       CASE #statRequest OF
         1:
           #data.parameterPage0 := #statParameterPage0;
         2:
           #data.systemCommand := #statSystemCommand;
         10:
           #data.vendorName := #statVendorName;
         11:
           #data.vendorText := #statVendorText;
         12:
           #data.productName := #statProductName;
         13:
           #data.productID := #statProductID;
         17:
           #data.fwRevision := #statFWRevision;
         18:
           #data.appSpecificName := #statAppSpecName;
         20:
           #data.statistics := #statStatistics;
         23:
           #data.diagnostics := #statDiagnostics;
         27:
           #data.parameters := #statParameters;
         ELSE // all other data sets are not defined
           ;
       END_CASE;
     END_IF;

     #statDone := #instDevice.done;
   END_REGION

   REGION OUTPUTS
     #done := #instDevice.done;
     #busy := #instDevice.busy;
     #error := #instDevice.error;
     #status := #instDevice.status;
     #diagDeviceFB := #instDevice.diagnostics;
   END_REGION
END_FUNCTION_BLOCK

// folder: Device-specific blocks/SIRIUS/3UG48

FUNCTION_BLOCK "LIOLink_3UG481x"   // FB5140, SCL
TITLE = LIOLink_3UG481x / IO_LINK_3UG481x
{ S7_Optimized_Access := 'FALSE' }
AUTHOR : SIOS
FAMILY : LIOLink
VERSION : 3.0
// IO-Link Device FB for SIRIUS 3UG481x to use with S7-300/400 controllers! / IO-Link Geraete FB fuer SIRIUS 3UG481x zur Nutzung mit S7-1500!
   VAR_INPUT
      execute : Bool;   // Request to execute function / Auftrag starten (mit steigender Flanke)
      logicalAddr : DInt;   // Logical address of IO-Link master module (sub module for ET 200eco PN) / Logische EA-Adresse des IO-Link Master Moduls
      cap : Int := 227;   // Client Access Point; 0xB400 for ET 200eco PN, CM 8x IO-Link, else 0xE003 (227) / Client Access Point (CAP), Siemens IO-Link Master immer 227 dezimal
      readWrite : Bool;   // FALSE: read, TRUE: write / Lese-/Schreibzugriff: 0=Lesen, 1=Schreiben
      port : Int;   // Port of the IO-Link Master for the Device / Port des Geraetes am IO-Link Mastermodul
      parameterPage0 : Bool := FALSE;   // Read access on parameter page 0 / Lesen Parameter Page 0
      systemCommands : Bool := FALSE;   // Write system commands / Schreiben Systemkommandos
      vendorName : Bool := FALSE;   // Read vendor name / Lesen Herstellername
      vendorText : Bool := FALSE;   // Read vendor text / Lesen Herstellertext
      productName : Bool := FALSE;   // Read product name / Lesen Produktname
      productID : Bool := FALSE;   // Read product ID / Lesen Produkt ID
      hwRevision : Bool := FALSE;   // Read hardware revision / Lesen HW-Revision
      fwRevision : Bool := FALSE;   // Read firmware revision / Lesen FW-Revision
      appSpecificName : Bool := FALSE;   // Read/Write application specific name / Lesen/Schreiben des spezifischen Applikationsnamen
      diagnostics : Bool := FALSE;   // Read diagnostics / Lesen der Diagnose
      measurements : Bool := FALSE;   // Read measurements / Lesen der Messwerte
      parameters : Bool;   // Read/Write parameters / Lesen/Schreiben der Parameter
   END_VAR
   VAR_OUTPUT
      done : Bool;   // TRUE: Commanded functionality has been completed successfully / Gueltigkeit 0: Daten ungueltig ; 1: Daten gueltig
      busy : Bool;   // TRUE: FB is not finished and new output values can be expected / 0: Auftrag beendet 1: Auftrag in Bearbeitung
      error : Bool;   // TRUE: An error occurred during the execution of the FB / Fehler = 0: kein Fehler; 1: Funktionsabbruch mit Fehler
      status : Word;   // 16#0000 - 16#7FFF: Status of the FB, 16#8000 - 16#FFFF: Error identification / DP/ PNIO - Fehlerstatus ; ERROR = 1 - Kommunikationsfehler in Detail
      diagDeviceFB : "LIOLink_typeDiagnostics";   // Diagnostics information of LIOLink_Device / IO-Link - Fehlerstatus; ERROR = 1: IO-Link Fehler in Detail
   END_VAR
   VAR_IN_OUT
      data : "LIOLink_3UG481_typeAll";   // Data area, device specific (Data Type) / Ablage der Gerätedaten, gerätespezifisch (Datentyp in DB)
   END_VAR
   VAR
      instDevice : "LIOLink_Device";
      statRecordParam : Struct   // Parameters to read/write specific records / Datensatzparameter (geraetespezifisch)
         index : Array[0..28] of Int;   // Index of data set / Datensatzindex
         subindex : Array[0..28] of Int;   // Subindex of data sets / Datensatzsubindex
         length : Array[0..28] of Int;   // Length of data set / Datensatzlänge
      END_STRUCT;
      statRecord : Array[0..231] of Byte;   // Record buffer
      statParameterPage0 AT statRecord : "LIOLink_typeParameterPage0";
      statSystemCommands AT statRecord : Byte;
      statVendorName AT statRecord : String[11];
      statVendorText AT statRecord : String[64];
      statProductName AT statRecord : String[64];
      statProductID AT statRecord : String[14];
      statHWRevision AT statRecord : String[7];
      statFWRevision AT statRecord : String[7];
      statAppSpecName AT statRecord : String[32];
      statDiagnostics AT statRecord : "LIOLink_3UG481_typeDiag";
      statMeasurements AT statRecord : "LIOLink_3UG481_typeMeasure";
      statParameters AT statRecord : "LIOLink_3UG481_typeParam";   // Product family SIRIUS (0x60)
      statIndex : Int;   // Requested index
      statSubindex : Int;   // Requested subindex
      statRecordLen : Int;   // Length of record to be written
      statRequest : Int;   // Case of request (data set) / Aktueller Fall (anfgefragter Datensatz)
      statDoneOld : Bool;   // Last cycle's value of instDevice.done
   END_VAR
   VAR_TEMP
      tempIndex : Int;   // Loop index
      tempLen : Int;   // Length
   END_VAR
   VAR CONSTANT
      MODE_READ : Bool := FALSE;   // Mode to read data
      MODE_WRITE : Bool := TRUE;   // Mode to write data
      STATUS_IDLE : Word := 16#7000;   // Status: Idle
   END_VAR
   // statRecordParam.index[3] := 2;
   // statRecordParam.index[2] := 0;
   // statRecordParam.index[1] := 0;
   // statRecordParam.index[0] := 0;
   // statRecordParam.index[17] := 23;
   // statRecordParam.index[16] := 22;
   // statRecordParam.index[5] := 0;
   // statRecordParam.index[4] := 0;
   // statRecordParam.index[15] := 21;
   // statRecordParam.index[14] := 20;
   // statRecordParam.index[13] := 19;
   // statRecordParam.index[12] := 18;
   // statRecordParam.index[11] := 17;
   // statRecordParam.index[10] := 16;
   // statRecordParam.index[9] := 0;
   // statRecordParam.index[8] := 0;
   // statRecordParam.index[7] := 0;
   // statRecordParam.index[6] := 0;
   // statRecordParam.length[28] := 60;
   // statRecordParam.length[27] := 0;
   // statRecordParam.length[26] := 0;
   // statRecordParam.length[25] := 38;
   // statRecordParam.length[24] := 30;
   // statRecordParam.length[23] := 0;
   // statRecordParam.length[22] := 0;
   // statRecordParam.length[21] := 0;
   // statRecordParam.length[20] := 0;
   // statRecordParam.length[19] := 0;
   // statRecordParam.length[18] := 32;
   // statRecordParam.length[17] := 7;
   // statRecordParam.length[16] := 7;
   // statRecordParam.length[15] := 0;
   // statRecordParam.length[14] := 0;
   // statRecordParam.length[13] := 14;
   // statRecordParam.length[12] := 64;
   // statRecordParam.length[11] := 64;
   // statRecordParam.length[10] := 11;
   // statRecordParam.length[9] := 0;
   // statRecordParam.length[8] := 0;
   // statRecordParam.length[7] := 0;
   // statRecordParam.length[6] := 0;
   // statRecordParam.length[5] := 0;
   // statRecordParam.length[4] := 0;
   // statRecordParam.length[3] := 1;
   // statRecordParam.length[2] := 0;
   // statRecordParam.length[1] := 16;
   // statRecordParam.length[0] := 0;
   // statRecordParam.index[28] := 131;
   // statRecordParam.index[27] := 0;
   // statRecordParam.index[26] := 0;
   // statRecordParam.index[25] := 94;
   // statRecordParam.index[24] := 92;
   // statRecordParam.index[23] := 0;
   // statRecordParam.index[22] := 0;
   // statRecordParam.index[21] := 0;
   // statRecordParam.index[20] := 0;
   // statRecordParam.index[19] := 0;
   // statRecordParam.index[18] := 24;
BEGIN
   REGION BLOCK INFO HEADER
     //===============================================================================
     // Siemens / (c)Copyright 2020
     //-------------------------------------------------------------------------------
     // Title:            LIOLink_3UG481x
     // Function:         Capsule block to communicate with 3UG481x devices
     // Library:          LIOLink
     // Author:           Siemens Industry Online Support
     // Tested with:      CPU 317-2 PN/DP FW 3.2
     // Engineering:      TIA Portal V16
     // Restrictions:     --
     // Requirements:     --
     //-------------------------------------------------------------------------------
     // Change log table:
     // Version  | Date       | Expert in charge       | Changes applied
     //----------|------------|------------------------|------------------------------
     // 01.00.00 | 11.04.2014 | Online Support         | First release
     // 01.01.00 | 12.09.2014 | Online Support         | Bugfixing write case 28 (data set 131)
     // 02.00.00 | 30.03.2015 | Online Support         | Upgrade to TIA Portal V13 SP1, use function IO_LINK_DEVICE, only one function for S7-1200 and 1500
     // 02.01.00 | 23.10.2015 | Online Support         | Upgraded FB "IO_LINK_DEVICE to V3.1.0
     // 03.00.00 | 22.09.2020 | Online Support         | Rewrote block for FB "LIOLink_Device" V4.0.0
     //===============================================================================
   END_REGION

   REGION INIT
     IF (#execute = TRUE AND #instDevice.status = #STATUS_IDLE) THEN
       // Request selector
       IF #parameterPage0 THEN
         #statRequest := 1;
       ELSIF #systemCommands THEN
         #statRequest := 3;
       ELSIF #vendorName THEN
         #statRequest := 10;
       ELSIF #vendorText THEN
         #statRequest := 11;
       ELSIF #productName THEN
         #statRequest := 12;
       ELSIF #productID THEN
         #statRequest := 13;
       ELSIF #hwRevision THEN
         #statRequest := 16;
       ELSIF #fwRevision THEN
         #statRequest := 17;
       ELSIF #appSpecificName THEN
         #statRequest := 18;
       ELSIF #diagnostics THEN
         #statRequest := 24;
       ELSIF #measurements THEN
         #statRequest := 25;
       ELSIF #parameters THEN
         #statRequest := 28;
       ELSE
         #statRequest := 0;
       END_IF;

       // Set request specific parameters
       #statIndex := #statRecordParam.index[#statRequest];
       #statSubindex := #statRecordParam.subindex[#statRequest];
       #statRecordLen := #statRecordParam.length[#statRequest];

       IF #readWrite = #MODE_WRITE THEN
         REGION write
           CASE #statRequest OF
             3:
               #statSystemCommands := #data.systemCommands;
             18:
               #statAppSpecName := #data.appSpecificName; // copy text into writing data
               #tempLen := LEN(#statAppSpecName); // determine length of text

               // Shift chars in array to remove String header
               FOR #tempIndex := 0 TO #tempLen - 1 DO
                 #statRecord[#tempIndex] := #statRecord[#tempIndex + 2]; // move [2] to [0], [3] to [1] ... until end of String
               END_FOR;

               // Fill remaining characters with null
               FOR #tempIndex := #tempLen TO #statRecordLen - 1 DO
                 #statRecord[#tempIndex] := CHAR_TO_BYTE('$00');
               END_FOR;
             28:
               #statParameters := #data.parameters;
             ELSE // All other data sets are read only  
               ;
           END_CASE;
         END_REGION

       END_IF;
     END_IF;
   END_REGION

   REGION CALL
     #instDevice(execute     := #execute,
                 logicalAddr := #logicalAddr,
                 cap         := #cap,
                 readWrite        := #readWrite,
                 "port"      := #port,
                 index       := #statIndex,
                 subindex    := #statSubindex,
                 writeLen    := #statRecordLen,
                 timeout     := T#20s,
                 record      := #statRecord);
   END_REGION

   REGION READ
     // Copy data
     IF #instDevice.done = TRUE AND #statDoneOld = FALSE AND #readWrite = #MODE_READ THEN
       IF (#statRequest >= 10 AND #statRequest <= 18) THEN // Only applies for String parameters (case 10..18)
         // Shift all characters to add string header
         FOR #tempIndex := (#statRecordLen + 1) TO 2 BY -1 DO
           #statRecord[#tempIndex] := #statRecord[#tempIndex - 2];
         END_FOR;
         // Add String header
         #statRecord[0] := INT_TO_BYTE(#statRecordLen);
         #statRecord[1] := INT_TO_BYTE(#statRecordLen);
       END_IF;

       CASE #statRequest OF
         1:
           #data.parameterPage0 := #statParameterPage0;
         10:
           #data.vendorName := #statVendorName;
         11:
           #data.vendorText := #statVendorText;
         12:
           #data.productName := #statProductName;
         13:
           #data.productID := #statProductID;
         16:
           #data.hwRevision := #statHWRevision;
         17:
           #data.fwRevision := #statFWRevision;
         18:
           #data.appSpecificName := #statAppSpecName;
         24:
           #data.diagnostics := #statDiagnostics;
         25:
           #data.measuredValues := #statMeasurements;
         28:
           #data.parameters := #statParameters;
         ELSE // Other data sets are not defined
           ;
       END_CASE;
     END_IF;

     #statDoneOld := #instDevice.done;
   END_REGION

   REGION OUTPUTS
     #done := #instDevice.done;
     #busy := #instDevice.busy;
     #error := #instDevice.error;
     #status := #instDevice.status;
     #diagDeviceFB := #instDevice.diagnostics;
   END_REGION
END_FUNCTION_BLOCK

FUNCTION_BLOCK "LIOLink_3UG4822"   // FB5150, SCL
TITLE = LIOLink_3UG4822 / IO_LINK_3UG4822_1500
{ S7_Optimized_Access := 'FALSE' }
AUTHOR : SIOS
FAMILY : LIOLink
VERSION : 3.0
// IO-Link Device FB for SIRIUS 3UG4822 to use with S7-300/400 controllers! / IO-Link Geraete FB fuer SIRIUS 3UG4822 zur Nutzung mit S7-1500!
   VAR_INPUT
      execute : Bool;   // Request to execute function / Auftrag starten (mit steigender Flanke)
      logicalAddr : DInt;   // Logical address of IO-Link master module (sub module for ET 200eco PN) / Logische EA-Adresse des IO-Link Master Moduls
      cap : Int := 227;   // Client Access Point; 0xB400 for ET 200eco PN, CM 8x IO-Link, else 0xE003 (227) / Client Access Point (CAP), Siemens IO-Link Master immer 227 dezimal
      readWrite : Bool;   // FALSE: read, TRUE: write / Lese-/Schreibzugriff: 0=Lesen, 1=Schreiben
      port : Int;   // Port of the IO-Link Master for the Device / Port des Geraetes am IO-Link Mastermodul
      parameterPage0 : Bool;   // Read access on parameter page 0 / Lesen Parameter Page 0
      systemCommands : Bool;   // Write system commands / Schreiben Systemkommandos
      vendorName : Bool;   // Read vendor name / Lesen Herstellername
      vendorText : Bool;   // Read vendor text / Lesen Herstellertext
      productName : Bool;   // Read product name / Lesen Produktname
      productID : Bool;   // Read product ID / Lesen Produkt ID
      hwRevision : Bool;   // Read hardware revision / Lesen HW-Revision
      fwRevision : Bool;   // Read firmware revision / Lesen FW-Revision
      appSpecificName : Bool;   // Read/Write application specific name / Lesen/Schreiben des spezifischen Applikationsnamen
      diagnostics : Bool;   // Read diagnostics / Lesen der Diagnose
      measurements : Bool;   // Read measurements / Lesen der Messwerte
      parameters : Bool;   // Read/Write parameters / Lesen/Schreiben der Parameter
   END_VAR
   VAR_OUTPUT
      done : Bool;   // TRUE: Commanded functionality has been completed successfully / Gueltigkeit 0: Daten ungueltig ; 1: Daten gueltig
      busy : Bool;   // TRUE: FB is not finished and new output values can be expected / 0: Auftrag beendet 1: Auftrag in Bearbeitung
      error : Bool;   // TRUE: An error occurred during the execution of the FB / Fehler = 0: kein Fehler; 1: Funktionsabbruch mit Fehler
      status : Word;   // 16#0000 - 16#7FFF: Status of the FB, 16#8000 - 16#FFFF: Error identification / DP/ PNIO - Fehlerstatus ; ERROR = 1 - Kommunikationsfehler in Detail
      diagDeviceFB : "LIOLink_typeDiagnostics";   // Diagnostics information of LIOLink_Device / IO-Link - Fehlerstatus; ERROR = 1: IO-Link Fehler in Detail
   END_VAR
   VAR_IN_OUT
      data : "LIOLink_3UG4822_typeAll";   // Data area, device specific (Data Type) / Ablage der Gerätedaten, gerätespezifisch (Datentyp in DB)
   END_VAR
   VAR
      instDevice : "LIOLink_Device";
      statRecordParam : Struct   // Parameters to read/write specific records / Datensatzparameter (geraetespezifisch)
         index : Array[0..28] of Int;   // Index of data set / Datensatzindex
         subindex : Array[0..28] of Int;   // Subindex of data sets / Datensatzsubindex
         length : Array[0..28] of Int;   // Length of data set / Datensatzlänge
      END_STRUCT;
      statRecord : Array[0..231] of Byte;   // Record buffer
      statParameterPage0 AT statRecord : "LIOLink_typeParameterPage0";
      statVendorName AT statRecord : String[11];
      statVendorText AT statRecord : String[64];
      statProductName AT statRecord : String[64];
      statProductID AT statRecord : String[14];
      statHWRevision AT statRecord : String[7];
      statFWRevision AT statRecord : String[7];
      statAppSpecName AT statRecord : String[32];
      statDiagnostics AT statRecord : "LIOLink_3UG4822_typeDiag";
      statMeasurements AT statRecord : "LIOLink_3UG4822_typeMeasure";
      statParameters AT statRecord : "LIOLink_3UG4822_typeParam";   // Product family SIRIUS (0x60)
      statSystemCommands AT statRecord : Byte;
      statIndex : Int;   // Requested index
      statSubindex : Int;   // Requested subindex
      statRecordLen : Int;   // Length of record to be written
      statRequest : Int;   // Case of request (data set) / Aktueller Fall (anfgefragter Datensatz)
      statDoneOld : Bool;   // Last cycle's value of instDevice.done
   END_VAR
   VAR_TEMP
      tempIndex : Int;   // Loop index
      tempLen : Int;   // Length
   END_VAR
   VAR CONSTANT
      MODE_READ : Bool := FALSE;   // Mode to read data
      MODE_WRITE : Bool := TRUE;   // Mode to write data
      STATUS_IDLE : Word := 16#7000;   // Status: Idle
   END_VAR
   // statRecordParam.index[3] := 2;
   // statRecordParam.index[2] := 0;
   // statRecordParam.index[1] := 0;
   // statRecordParam.index[0] := 0;
   // statRecordParam.index[17] := 23;
   // statRecordParam.index[16] := 22;
   // statRecordParam.index[5] := 0;
   // statRecordParam.index[4] := 0;
   // statRecordParam.index[15] := 21;
   // statRecordParam.index[14] := 20;
   // statRecordParam.index[13] := 19;
   // statRecordParam.index[12] := 18;
   // statRecordParam.index[11] := 17;
   // statRecordParam.index[10] := 16;
   // statRecordParam.index[9] := 0;
   // statRecordParam.index[8] := 0;
   // statRecordParam.index[7] := 0;
   // statRecordParam.index[6] := 0;
   // statRecordParam.length[28] := 64;
   // statRecordParam.length[27] := 0;
   // statRecordParam.length[26] := 0;
   // statRecordParam.length[25] := 52;
   // statRecordParam.length[24] := 28;
   // statRecordParam.length[23] := 0;
   // statRecordParam.length[22] := 0;
   // statRecordParam.length[21] := 0;
   // statRecordParam.length[20] := 0;
   // statRecordParam.length[19] := 0;
   // statRecordParam.length[18] := 32;
   // statRecordParam.length[17] := 7;
   // statRecordParam.length[16] := 7;
   // statRecordParam.length[15] := 0;
   // statRecordParam.length[14] := 0;
   // statRecordParam.length[13] := 14;
   // statRecordParam.length[12] := 64;
   // statRecordParam.length[11] := 64;
   // statRecordParam.length[10] := 11;
   // statRecordParam.length[9] := 0;
   // statRecordParam.length[8] := 0;
   // statRecordParam.length[7] := 0;
   // statRecordParam.length[6] := 0;
   // statRecordParam.length[5] := 0;
   // statRecordParam.length[4] := 0;
   // statRecordParam.length[3] := 1;
   // statRecordParam.length[2] := 0;
   // statRecordParam.length[1] := 16;
   // statRecordParam.length[0] := 0;
   // statRecordParam.index[28] := 131;
   // statRecordParam.index[27] := 0;
   // statRecordParam.index[26] := 0;
   // statRecordParam.index[25] := 94;
   // statRecordParam.index[24] := 92;
   // statRecordParam.index[23] := 0;
   // statRecordParam.index[22] := 0;
   // statRecordParam.index[21] := 0;
   // statRecordParam.index[20] := 0;
   // statRecordParam.index[19] := 0;
   // statRecordParam.index[18] := 24;
BEGIN
   REGION BLOCK INFO HEADER
     //===============================================================================
     // Siemens / (c)Copyright 2020
     //-------------------------------------------------------------------------------
     // Title:            LIOLink_3UG4822
     // Function:         Capsule block to communicate with 3UG4822 devices
     // Library:          LIOLink
     // Author:           Siemens Industry Online Support
     // Tested with:      CPU 317-2 PN/DP FW 3.2
     // Engineering:      TIA Portal V16
     // Restrictions:     --
     // Requirements:     --
     //-------------------------------------------------------------------------------
     // Change log table:
     // Version  | Date       | Expert in charge       | Changes applied
     //----------|------------|------------------------|------------------------------
     // 01.00.00 | 11.04.2014 | Online Support         | First release
     // 01.01.00 | 12.09.2014 | Online Support         | Bugfixing write case 28 (data set 131)
     // 02.00.00 | 30.03.2015 | Online Support         | Upgrade to TIA Portal V13 SP1, use function IO_LINK_DEVICE, only one function for S7-1200 and 1500
     // 02.01.00 | 23.10.2015 | Online Support         | Upgraded FB "IO_LINK_DEVICE to V3.1.0
     // 03.00.00 | 22.09.2020 | Online Support         | Rewrote block for FB "LIOLink_Device" V4.0.0
     //===============================================================================
   END_REGION

   REGION INIT
     IF (#execute = TRUE AND #instDevice.status = #STATUS_IDLE) THEN
       // Request selector
       IF #parameterPage0 THEN
         #statRequest := 1;
       ELSIF #systemCommands THEN
         #statRequest := 3;
       ELSIF #vendorName THEN
         #statRequest := 10;
       ELSIF #vendorText THEN
         #statRequest := 11;
       ELSIF #productName THEN
         #statRequest := 12;
       ELSIF #productID THEN
         #statRequest := 13;
       ELSIF #hwRevision THEN
         #statRequest := 16;
       ELSIF #fwRevision THEN
         #statRequest := 17;
       ELSIF #appSpecificName THEN
         #statRequest := 18;
       ELSIF #diagnostics THEN
         #statRequest := 24;
       ELSIF #measurements THEN
         #statRequest := 25;
       ELSIF #parameters THEN
         #statRequest := 28;
       ELSE
         #statRequest := 0;
       END_IF;

       // Set request specific parameters
       #statIndex := #statRecordParam.index[#statRequest];
       #statSubindex := #statRecordParam.subindex[#statRequest];
       #statRecordLen := #statRecordParam.length[#statRequest];

       IF #readWrite = #MODE_WRITE THEN
         REGION write
           CASE #statRequest OF
             3:
               #statSystemCommands := #data.systemCommands;
             18:
               #statAppSpecName := #data.appSpecificName; // copy text into writing data
               #tempLen := LEN(#statAppSpecName); // determine length of text

               // Shift chars in array to remove String header
               FOR #tempIndex := 0 TO #tempLen - 1 DO
                 #statRecord[#tempIndex] := #statRecord[#tempIndex + 2]; // move [2] to [0], [3] to [1] ... until end of String
               END_FOR;

               // Fill remaining characters with null
               FOR #tempIndex := #tempLen TO #statRecordLen - 1 DO
                 #statRecord[#tempIndex] := CHAR_TO_BYTE('$00');
               END_FOR;
             28:
               #statParameters := #data.parameters;
             ELSE // All other data sets are read only  
               ;
           END_CASE;
         END_REGION

       END_IF;
     END_IF;
   END_REGION

   REGION CALL
     #instDevice(execute     := #execute,
                 logicalAddr := #logicalAddr,
                 cap         := #cap,
                 readWrite   := #readWrite,
                 "port"      := #port,
                 index       := #statIndex,
                 subindex    := #statSubindex,
                 writeLen    := #statRecordLen,
                 timeout     := T#20s,
                 record      := #statRecord);
   END_REGION

   REGION READ
     // Copy data
     IF #instDevice.done = TRUE AND #statDoneOld = FALSE AND #readWrite = #MODE_READ THEN
       IF (#statRequest >= 10 AND #statRequest <= 18) THEN // Only applies for String parameters (case 10..18)
         // Shift all characters to add string header
         FOR #tempIndex := (#statRecordLen + 1) TO 2 BY -1 DO
           #statRecord[#tempIndex] := #statRecord[#tempIndex - 2];
         END_FOR;
         // Add String header
         #statRecord[0] := INT_TO_BYTE(#statRecordLen);
         #statRecord[1] := INT_TO_BYTE(#statRecordLen);
       END_IF;

       CASE #statRequest OF
         1:
           #data.parameterPage0 := #statParameterPage0;
         10:
           #data.vendorName := #statVendorName;
         11:
           #data.vendorText := #statVendorText;
         12:
           #data.productName := #statProductName;
         13:
           #data.productID := #statProductID;
         16:
           #data.hwRevision := #statHWRevision;
         17:
           #data.fwRevision := #statFWRevision;
         18:
           #data.appSpecificName := #statAppSpecName;
         24:
           #data.diagnostics := #statDiagnostics;
         25:
           #data.measuredValues := #statMeasurements;
         28:
           #data.parameters := #statParameters;
         ELSE // Other data sets are not defined
           ;
       END_CASE;
     END_IF;

     #statDoneOld := #instDevice.done;
   END_REGION

   REGION OUTPUTS
     #done := #instDevice.done;
     #busy := #instDevice.busy;
     #error := #instDevice.error;
     #status := #instDevice.status;
     #diagDeviceFB := #instDevice.diagnostics;
   END_REGION
END_FUNCTION_BLOCK

FUNCTION_BLOCK "LIOLink_3UG4825"   // FB5160, SCL
TITLE = LIOLink_3UG4825 / IO_LINK_3UG4825_1500
{ S7_Optimized_Access := 'FALSE' }
AUTHOR : SIOS
FAMILY : LIOLink
VERSION : 3.0
// IO-Link Device FB for SIRIUS 3UG4825 to use with S7-300/400 controllers! / IO-Link Geraete FB fuer SIRIUS 3UG4825 zur Nutzung mit S7-1500!
   VAR_INPUT
      execute : Bool;   // Request to execute function / Auftrag starten (mit steigender Flanke)
      logicalAddr : DInt;   // Logical address of IO-Link master module (sub module for ET 200eco PN) / Logische EA-Adresse des IO-Link Master Moduls
      cap : Int := 227;   // Client Access Point; 0xB400 for ET 200eco PN, CM 8x IO-Link, else 0xE003 (227) / Client Access Point (CAP), Siemens IO-Link Master immer 227 dezimal
      readWrite : Bool;   // FALSE: read, TRUE: write / Lese-/Schreibzugriff: 0=Lesen, 1=Schreiben
      port : Int;   // Port of the IO-Link Master for the Device / Port des Geraetes am IO-Link Mastermodul
      parameterPage0 : Bool;   // Read access on parameter page 0 / Lesen Parameter Page 0
      systemCommands : Bool;   // Write system commands / Schreiben Systemkommandos
      vendorName : Bool;   // Read vendor name / Lesen Herstellername
      vendorText : Bool;   // Read vendor text / Lesen Herstellertext
      productName : Bool;   // Read product name / Lesen Produktname
      productID : Bool;   // Read product ID / Lesen Produkt ID
      serialNumber : Bool;   // Read serial number / Lesen Seriennummer
      hwRevision : Bool;   // Read hardware revision / Lesen HW-Revision
      fwRevision : Bool;   // Read firmware revision / Lesen FW-Revision
      appSpecificName : Bool;   // Read/Write application specific name / Lesen/Schreiben des spezifischen Applikationsnamen
      diagnostics : Bool;   // Read diagnostics / Lesen der Diagnose
      measurements : Bool;   // Read measurements / Lesen der Messwerte
      parameters : Bool;   // Read/Write parameters / Lesen/Schreiben der Parameter
   END_VAR
   VAR_OUTPUT
      done : Bool;   // TRUE: Commanded functionality has been completed successfully / Gueltigkeit 0: Daten ungueltig ; 1: Daten gueltig
      busy : Bool;   // TRUE: FB is not finished and new output values can be expected / 0: Auftrag beendet 1: Auftrag in Bearbeitung
      error : Bool;   // TRUE: An error occurred during the execution of the FB / Fehler = 0: kein Fehler; 1: Funktionsabbruch mit Fehler
      status : Word;   // 16#0000 - 16#7FFF: Status of the FB, 16#8000 - 16#FFFF: Error identification / DP/ PNIO - Fehlerstatus ; ERROR = 1 - Kommunikationsfehler in Detail
      diagDeviceFB : "LIOLink_typeDiagnostics";   // Diagnostics information of LIOLink_Device / IO-Link - Fehlerstatus; ERROR = 1: IO-Link Fehler in Detail
   END_VAR
   VAR_IN_OUT
      data : "LIOLink_3UG4825_typeAll";   // Data area, device specific (Data Type) / Ablage der Gerätedaten, gerätespezifisch (Datentyp in DB)
   END_VAR
   VAR
      instDevice : "LIOLink_Device";
      statRecordParam : Struct   // Parameters to read/write specific records / Datensatzparameter (geraetespezifisch)
         index : Array[0..28] of Int;   // Index of data set / Datensatzindex
         subindex : Array[0..28] of Int;   // Subindex of data sets / Datensatzsubindex
         length : Array[0..28] of Int;   // Length of data set / Datensatzlänge
      END_STRUCT;
      statRecord : Array[0..231] of Byte;   // Record buffer
      statParameterPage0 AT statRecord : "LIOLink_typeParameterPage0";
      statVendorName AT statRecord : String[11];
      statVendorText AT statRecord : String[64];
      statProductName AT statRecord : String[64];
      statProductID AT statRecord : String[14];
      statSerialNumber AT statRecord : String[16];
      statHWRevision AT statRecord : String[7];
      statFWRevision AT statRecord : String[7];
      statAppSpecName AT statRecord : String[32];
      statDiagnostics AT statRecord : "LIOLink_3UG4825_typeDiag";
      statMeasurements AT statRecord : "LIOLink_3UG4825_typeMeasure";
      statParameters AT statRecord : "LIOLink_3UG4825_typeParam";   // Product family SIRIUS (0x60)
      statSystemCommands AT statRecord : Byte;
      statIndex : Int;   // Requested index
      statSubindex : Int;   // Requested subindex
      statRecordLen : Int;   // Length of record to be written
      statRequest : Int;   // Case of request (data set) / Aktueller Fall (anfgefragter Datensatz)
      statDoneOld : Bool;   // Last cycle's value of instDevice.done
   END_VAR
   VAR_TEMP
      tempIndex : Int;   // Loop index
      tempLen : Int;   // Length
   END_VAR
   VAR CONSTANT
      MODE_READ : Bool := FALSE;   // Mode to read data
      MODE_WRITE : Bool := TRUE;   // Mode to write data
      STATUS_IDLE : Word := 16#7000;   // Status: Idle
   END_VAR
   // statRecordParam.index[3] := 2;
   // statRecordParam.index[2] := 0;
   // statRecordParam.index[1] := 0;
   // statRecordParam.index[0] := 0;
   // statRecordParam.index[18] := 24;
   // statRecordParam.index[17] := 23;
   // statRecordParam.index[5] := 0;
   // statRecordParam.index[4] := 0;
   // statRecordParam.index[16] := 22;
   // statRecordParam.index[15] := 21;
   // statRecordParam.index[14] := 20;
   // statRecordParam.index[13] := 19;
   // statRecordParam.index[12] := 18;
   // statRecordParam.index[11] := 17;
   // statRecordParam.index[10] := 16;
   // statRecordParam.index[9] := 0;
   // statRecordParam.index[8] := 0;
   // statRecordParam.index[7] := 0;
   // statRecordParam.index[6] := 0;
   // statRecordParam.length[28] := 48;
   // statRecordParam.length[27] := 0;
   // statRecordParam.length[26] := 0;
   // statRecordParam.length[25] := 22;
   // statRecordParam.length[24] := 30;
   // statRecordParam.length[23] := 0;
   // statRecordParam.length[22] := 0;
   // statRecordParam.length[21] := 0;
   // statRecordParam.length[20] := 0;
   // statRecordParam.length[19] := 0;
   // statRecordParam.length[18] := 32;
   // statRecordParam.length[17] := 7;
   // statRecordParam.length[16] := 7;
   // statRecordParam.length[15] := 16;
   // statRecordParam.length[14] := 0;
   // statRecordParam.length[13] := 14;
   // statRecordParam.length[12] := 64;
   // statRecordParam.length[11] := 64;
   // statRecordParam.length[10] := 11;
   // statRecordParam.length[9] := 0;
   // statRecordParam.length[8] := 0;
   // statRecordParam.length[7] := 0;
   // statRecordParam.length[6] := 0;
   // statRecordParam.length[5] := 0;
   // statRecordParam.length[4] := 0;
   // statRecordParam.length[3] := 1;
   // statRecordParam.length[2] := 0;
   // statRecordParam.length[1] := 16;
   // statRecordParam.length[0] := 0;
   // statRecordParam.index[28] := 131;
   // statRecordParam.index[27] := 0;
   // statRecordParam.index[26] := 0;
   // statRecordParam.index[25] := 94;
   // statRecordParam.index[24] := 92;
   // statRecordParam.index[23] := 0;
   // statRecordParam.index[22] := 0;
   // statRecordParam.index[21] := 0;
   // statRecordParam.index[20] := 0;
   // statRecordParam.index[19] := 0;
BEGIN
   REGION BLOCK INFO HEADER
     //===============================================================================
     // Siemens / (c)Copyright 2020
     //-------------------------------------------------------------------------------
     // Title:            LIOLink_3UG4825
     // Function:         Capsule block to communicate with 3UG4825 devices
     // Library:          LIOLink
     // Author:           Siemens Industry Online Support
     // Tested with:      CPU 317-2 PN/DP FW 3.2
     // Engineering:      TIA Portal V16
     // Restrictions:     --
     // Requirements:     --
     //------------------------------------------------------------------------------
     // Change log table:
     // Version  | Date       | Expert in charge       | Changes applied
     //----------|------------|------------------------|------------------------------
     // 01.00.00 | 11.04.2014 | Online Support         | First release
     // 01.01.00 | 12.09.2014 | Online Support         | Bugfixing write case 28 (data set 131)
     // 02.00.00 | 30.03.2015 | Online Support         | Upgrade to TIA Portal V13 SP1, use function IO_LINK_DEVICE, only one function for S7-1200 and 1500
     // 02.01.00 | 23.10.2015 | Online Support         | Upgraded FB "IO_LINK_DEVICE to V3.1.0
     // 03.00.00 | 22.09.2020 | Online Support         | Rewrote block for FB "LIOLink_Device" V4.0.0
     //===============================================================================
   END_REGION

   REGION INIT
     IF (#execute = TRUE AND #instDevice.status = #STATUS_IDLE) THEN
       // Request selector
       IF #parameterPage0 THEN
         #statRequest := 1;
       ELSIF #systemCommands THEN
         #statRequest := 3;
       ELSIF #vendorName THEN
         #statRequest := 10;
       ELSIF #vendorText THEN
         #statRequest := 11;
       ELSIF #productName THEN
         #statRequest := 12;
       ELSIF #productID THEN
         #statRequest := 13;
       ELSIF #hwRevision THEN
         #statRequest := 16;
       ELSIF #fwRevision THEN
         #statRequest := 17;
       ELSIF #appSpecificName THEN
         #statRequest := 18;
       ELSIF #diagnostics THEN
         #statRequest := 24;
       ELSIF #measurements THEN
         #statRequest := 25;
       ELSIF #parameters THEN
         #statRequest := 28;
       ELSE
         #statRequest := 0;
       END_IF;

       // Set request specific parameters
       #statIndex := #statRecordParam.index[#statRequest];
       #statSubindex := #statRecordParam.subindex[#statRequest];
       #statRecordLen := #statRecordParam.length[#statRequest];

       IF #readWrite = #MODE_WRITE THEN
         REGION write
           CASE #statRequest OF
             3:
               #statSystemCommands := #data.systemCommands;
             18:
               #statAppSpecName := #data.appSpecificName; // copy text into writing data
               #tempLen := LEN(#statAppSpecName); // determine length of text

               // Shift chars in array to remove String header
               FOR #tempIndex := 0 TO #tempLen - 1 DO
                 #statRecord[#tempIndex] := #statRecord[#tempIndex + 2]; // move [2] to [0], [3] to [1] ... until end of String
               END_FOR;

               // Fill remaining characters with null
               FOR #tempIndex := #tempLen TO #statRecordLen - 1 DO
                 #statRecord[#tempIndex] := CHAR_TO_BYTE('$00');
               END_FOR;
             28:
               #statParameters := #data.parameters;
             ELSE // All other data sets are read only  
               ;
           END_CASE;
         END_REGION

       END_IF;
     END_IF;
   END_REGION

   REGION CALL
     #instDevice(execute     := #execute,
                 logicalAddr := #logicalAddr,
                 cap         := #cap,
                 readWrite   := #readWrite,
                 "port"      := #port,
                 index       := #statIndex,
                 subindex    := #statSubindex,
                 writeLen    := #statRecordLen,
                 timeout     := T#20s,
                 record      := #statRecord);
   END_REGION

   REGION READ
     // Copy data
     IF #instDevice.done = TRUE AND #statDoneOld = FALSE AND #readWrite = #MODE_READ THEN
       IF (#statRequest >= 10 AND #statRequest <= 18) THEN // Only applies for String parameters (case 10..18)
         // Shift all characters to add string header
         FOR #tempIndex := (#statRecordLen + 1) TO 2 BY -1 DO
           #statRecord[#tempIndex] := #statRecord[#tempIndex - 2];
         END_FOR;
         // Add String header
         #statRecord[0] := INT_TO_BYTE(#statRecordLen);
         #statRecord[1] := INT_TO_BYTE(#statRecordLen);
       END_IF;

       CASE #statRequest OF
         1:
           #data.parameterPage0 := #statParameterPage0;
         10:
           #data.vendorName := #statVendorName;
         11:
           #data.vendorText := #statVendorText;
         12:
           #data.productName := #statProductName;
         13:
           #data.productID := #statProductID;
         16:
           #data.hwRevision := #statHWRevision;
         17:
           #data.fwRevision := #statFWRevision;
         18:
           #data.appSpecificName := #statAppSpecName;
         24:
           #data.diagnostics := #statDiagnostics;
         25:
           #data.measuredValues := #statMeasurements;
         28:
           #data.parameters := #statParameters;
         ELSE // Other data sets are not defined
           ;
       END_CASE;
     END_IF;

     #statDoneOld := #instDevice.done;
   END_REGION

   REGION OUTPUTS
     #done := #instDevice.done;
     #busy := #instDevice.busy;
     #error := #instDevice.error;
     #status := #instDevice.status;
     #diagDeviceFB := #instDevice.diagnostics;
   END_REGION
END_FUNCTION_BLOCK

FUNCTION_BLOCK "LIOLink_3UG4832"   // FB5170, SCL
TITLE = LIOLink_3UG4832 / IO_LINK_3UG4832_1500
{ S7_Optimized_Access := 'FALSE' }
AUTHOR : SIOS
FAMILY : LIOLink
VERSION : 3.0
// IO-Link Device FB for SIRIUS 3UG4832 to use with S7-300/400 controllers! / IO-Link Geraete FB fuer SIRIUS 3UG4832 zur Nutzung mit S7-1500!
   VAR_INPUT
      execute : Bool;   // Request to execute function / Auftrag starten (mit steigender Flanke)
      logicalAddr : DInt;   // Logical address of IO-Link master module (sub module for ET 200eco PN) / Logische EA-Adresse des IO-Link Master Moduls
      cap : Int := 227;   // Client Access Point; 0xB400 for ET 200eco PN, CM 8x IO-Link, else 0xE003 (227) / Client Access Point (CAP), Siemens IO-Link Master immer 227 dezimal
      readWrite : Bool;   // FALSE: read, TRUE: write / Lese-/Schreibzugriff: 0=Lesen, 1=Schreiben
      port : Int;   // Port of the IO-Link Master for the Device / Port des Geraetes am IO-Link Mastermodul
      parameterPage0 : Bool;   // Read access on parameter page 0 / Lesen Parameter Page 0
      systemCommands : Bool;   // Write system commands / Schreiben Systemkommandos
      vendorName : Bool;   // Read vendor name / Lesen Herstellername
      vendorText : Bool;   // Read vendor text / Lesen Herstellertext
      productName : Bool;   // Read product name / Lesen Produktname
      productID : Bool;   // Read product ID / Lesen Produkt ID
      hwRevision : Bool;   // Read hardware revision / Lesen HW-Revision
      fwRevision : Bool;   // Read firmware revision / Lesen FW-Revision
      appSpecificName : Bool;   // Read/Write application specific name / Lesen/Schreiben des spezifischen Applikationsnamen
      diagnostics : Bool;   // Read diagnostics / Lesen der Diagnose
      measurements : Bool;   // Read measurements / Lesen der Messwerte
      parameters : Bool;   // Read/Write parameters / Lesen/Schreiben der Parameter
   END_VAR
   VAR_OUTPUT
      done : Bool;   // TRUE: Commanded functionality has been completed successfully / Gueltigkeit 0: Daten ungueltig ; 1: Daten gueltig
      busy : Bool;   // TRUE: FB is not finished and new output values can be expected / 0: Auftrag beendet 1: Auftrag in Bearbeitung
      error : Bool;   // TRUE: An error occurred during the execution of the FB / Fehler = 0: kein Fehler; 1: Funktionsabbruch mit Fehler
      status : Word;   // 16#0000 - 16#7FFF: Status of the FB, 16#8000 - 16#FFFF: Error identification / DP/ PNIO - Fehlerstatus ; ERROR = 1 - Kommunikationsfehler in Detail
      diagDeviceFB : "LIOLink_typeDiagnostics";   // Diagnostics information of LIOLink_Device / IO-Link - Fehlerstatus; ERROR = 1: IO-Link Fehler in Detail
   END_VAR
   VAR_IN_OUT
      data : "LIOLink_3UG4832_typeAll";   // Data area, device specific (Data Type) / Ablage der Gerätedaten, gerätespezifisch (Datentyp in DB)
   END_VAR
   VAR
      instDevice : "LIOLink_Device";
      statRecordParam : Struct   // Parameters to read/write specific records / Datensatzparameter (geraetespezifisch)
         index : Array[0..28] of Int;   // Index of data set / Datensatzindex
         subindex : Array[0..28] of Int;   // Subindex of data sets / Datensatzsubindex
         length : Array[0..28] of Int;   // Length of data set / Datensatzlänge
      END_STRUCT;
      statRecord : Array[0..231] of Byte;   // Record buffer
      statParameterPage0 AT statRecord : "LIOLink_typeParameterPage0";
      statVendorName AT statRecord : String[11];
      statVendorText AT statRecord : String[64];
      statProductName AT statRecord : String[64];
      statProductID AT statRecord : String[14];
      statHWRevision AT statRecord : String[7];
      statFWRevision AT statRecord : String[7];
      statAppSpecName AT statRecord : String[32];
      statDiagnostics AT statRecord : "LIOLink_3UG4832_typeDiag";
      statMeasurements AT statRecord : "LIOLink_3UG4832_typeMeasure";
      statParameters AT statRecord : "LIOLink_3UG4832_typeParam";   // Product family SIRIUS (0x60)
      statSystemCommands AT statRecord : Byte;
      statIndex : Int;   // Requested index
      statSubindex : Int;   // Requested subindex
      statRecordLen : Int;   // Length of record to be written
      statRequest : Int;   // Case of request (data set) / Aktueller Fall (anfgefragter Datensatz)
      statDoneOld : Bool;   // Last cycle's value of instDevice.done
   END_VAR
   VAR_TEMP
      tempIndex : Int;   // Loop index
      tempLen : Int;   // Length
   END_VAR
   VAR CONSTANT
      MODE_READ : Bool := FALSE;   // Mode to read data
      MODE_WRITE : Bool := TRUE;   // Mode to write data
      STATUS_IDLE : Word := 16#7000;   // Status: Idle
   END_VAR
   // statRecordParam.index[3] := 2;
   // statRecordParam.index[2] := 0;
   // statRecordParam.index[1] := 0;
   // statRecordParam.index[0] := 0;
   // statRecordParam.index[17] := 23;
   // statRecordParam.index[16] := 22;
   // statRecordParam.index[5] := 0;
   // statRecordParam.index[4] := 0;
   // statRecordParam.index[15] := 21;
   // statRecordParam.index[14] := 20;
   // statRecordParam.index[13] := 19;
   // statRecordParam.index[12] := 18;
   // statRecordParam.index[11] := 17;
   // statRecordParam.index[10] := 16;
   // statRecordParam.index[9] := 0;
   // statRecordParam.index[8] := 0;
   // statRecordParam.index[7] := 0;
   // statRecordParam.index[6] := 0;
   // statRecordParam.length[28] := 48;
   // statRecordParam.length[27] := 0;
   // statRecordParam.length[26] := 0;
   // statRecordParam.length[25] := 28;
   // statRecordParam.length[24] := 28;
   // statRecordParam.length[23] := 0;
   // statRecordParam.length[22] := 0;
   // statRecordParam.length[21] := 0;
   // statRecordParam.length[20] := 0;
   // statRecordParam.length[19] := 0;
   // statRecordParam.length[18] := 32;
   // statRecordParam.length[17] := 7;
   // statRecordParam.length[16] := 7;
   // statRecordParam.length[15] := 0;
   // statRecordParam.length[14] := 0;
   // statRecordParam.length[13] := 14;
   // statRecordParam.length[12] := 64;
   // statRecordParam.length[11] := 64;
   // statRecordParam.length[10] := 11;
   // statRecordParam.length[9] := 0;
   // statRecordParam.length[8] := 0;
   // statRecordParam.length[7] := 0;
   // statRecordParam.length[6] := 0;
   // statRecordParam.length[5] := 0;
   // statRecordParam.length[4] := 0;
   // statRecordParam.length[3] := 1;
   // statRecordParam.length[2] := 0;
   // statRecordParam.length[1] := 16;
   // statRecordParam.length[0] := 0;
   // statRecordParam.index[28] := 131;
   // statRecordParam.index[27] := 0;
   // statRecordParam.index[26] := 0;
   // statRecordParam.index[25] := 94;
   // statRecordParam.index[24] := 92;
   // statRecordParam.index[23] := 0;
   // statRecordParam.index[22] := 0;
   // statRecordParam.index[21] := 0;
   // statRecordParam.index[20] := 0;
   // statRecordParam.index[19] := 0;
   // statRecordParam.index[18] := 24;
BEGIN
   REGION BLOCK INFO HEADER
     //===============================================================================
     // Siemens / (c)Copyright 2020
     //-------------------------------------------------------------------------------
     // Title:            LIOLink_3UG4832
     // Function:         Capsule block to communicate with 3UG4832 devices
     // Library:          LIOLink
     // Author:           Siemens Industry Online Support
     // Tested with:      CPU 317-2 PN/DP FW 3.2
     // Engineering:      TIA Portal V16
     // Restrictions:     --
     // Requirements:     --
     //-------------------------------------------------------------------------------
     // Change log table:
     // Version  | Date       | Expert in charge       | Changes applied
     //----------|------------|------------------------|------------------------------
     // 01.00.00 | 11.04.2014 | Online Support         | First release
     // 01.01.00 | 12.09.2014 | Online Support         | Bugfixing write case 28 (data set 131)
     // 02.00.00 | 30.03.2015 | Online Support         | Upgrade to TIA Portal V13 SP1, use function IO_LINK_DEVICE, only one function for S7-1200 and 1500
     // 02.01.00 | 23.10.2015 | Online Support         | Upgraded FB "IO_LINK_DEVICE to V3.1.0
     // 03.00.00 | 22.09.2020 | Online Support         | Rewrote block for FB "LIOLink_Device" V4.0.0
     //===============================================================================
   END_REGION

   REGION INIT
     IF (#execute = TRUE AND #instDevice.status = #STATUS_IDLE) THEN
       // Request selector
       IF #parameterPage0 THEN
         #statRequest := 1;
       ELSIF #systemCommands THEN
         #statRequest := 3;
       ELSIF #vendorName THEN
         #statRequest := 10;
       ELSIF #vendorText THEN
         #statRequest := 11;
       ELSIF #productName THEN
         #statRequest := 12;
       ELSIF #productID THEN
         #statRequest := 13;
       ELSIF #hwRevision THEN
         #statRequest := 16;
       ELSIF #fwRevision THEN
         #statRequest := 17;
       ELSIF #appSpecificName THEN
         #statRequest := 18;
       ELSIF #diagnostics THEN
         #statRequest := 24;
       ELSIF #measurements THEN
         #statRequest := 25;
       ELSIF #parameters THEN
         #statRequest := 28;
       ELSE
         #statRequest := 0;
       END_IF;

       // Set request specific parameters
       #statIndex := #statRecordParam.index[#statRequest];
       #statSubindex := #statRecordParam.subindex[#statRequest];
       #statRecordLen := #statRecordParam.length[#statRequest];

       IF #readWrite = #MODE_WRITE THEN
         REGION write
           CASE #statRequest OF
             3:
               #statSystemCommands := #data.systemCommands;
             18:
               #statAppSpecName := #data.appSpecificName; // copy text into writing data
               #tempLen := LEN(#statAppSpecName); // determine length of text

               // Shift chars in array to remove String header
               FOR #tempIndex := 0 TO #tempLen - 1 DO
                 #statRecord[#tempIndex] := #statRecord[#tempIndex + 2]; // move [2] to [0], [3] to [1] ... until end of String
               END_FOR;

               // Fill remaining characters with null
               FOR #tempIndex := #tempLen TO #statRecordLen - 1 DO
                 #statRecord[#tempIndex] := CHAR_TO_BYTE('$00');
               END_FOR;
             28:
               #statParameters := #data.parameters;
             ELSE // All other data sets are read only  
               ;
           END_CASE;
         END_REGION

       END_IF;
     END_IF;
   END_REGION

   REGION CALL
     #instDevice(execute     := #execute,
                 logicalAddr := #logicalAddr,
                 cap         := #cap,
                 readWrite   := #readWrite,
                 "port"      := #port,
                 index       := #statIndex,
                 subindex    := #statSubindex,
                 writeLen    := #statRecordLen,
                 timeout     := T#20s,
                 record      := #statRecord);
   END_REGION

   REGION READ
     // Copy data
     IF #instDevice.done = TRUE AND #statDoneOld = FALSE AND #readWrite = #MODE_READ THEN
       IF (#statRequest >= 10 AND #statRequest <= 18) THEN // Only applies for String parameters (case 10..18)
         // Shift all characters to add string header
         FOR #tempIndex := (#statRecordLen + 1) TO 2 BY -1 DO
           #statRecord[#tempIndex] := #statRecord[#tempIndex - 2];
         END_FOR;
         // Add String header
         #statRecord[0] := INT_TO_BYTE(#statRecordLen);
         #statRecord[1] := INT_TO_BYTE(#statRecordLen);
       END_IF;

       CASE #statRequest OF
         1:
           #data.parameterPage0 := #statParameterPage0;
         10:
           #data.vendorName := #statVendorName;
         11:
           #data.vendorText := #statVendorText;
         12:
           #data.productName := #statProductName;
         13:
           #data.productID := #statProductID;
         16:
           #data.hwRevision := #statHWRevision;
         17:
           #data.fwRevision := #statFWRevision;
         18:
           #data.appSpecificName := #statAppSpecName;
         24:
           #data.diagnostics := #statDiagnostics;
         25:
           #data.measuredValues := #statMeasurements;
         28:
           #data.parameters := #statParameters;
         ELSE // Other data sets are not defined
           ;
       END_CASE;
     END_IF;

     #statDoneOld := #instDevice.done;
   END_REGION

   REGION OUTPUTS
     #done := #instDevice.done;
     #busy := #instDevice.busy;
     #error := #instDevice.error;
     #status := #instDevice.status;
     #diagDeviceFB := #instDevice.diagnostics;
   END_REGION
END_FUNCTION_BLOCK

FUNCTION_BLOCK "LIOLink_3UG4841"   // FB5180, SCL
TITLE = LIOLink_3UG4841 / IO_LINK_3UG4841_1500
{ S7_Optimized_Access := 'FALSE' }
AUTHOR : SIOS
FAMILY : LIOLink
VERSION : 3.0
// IO-Link Device FB for SIRIUS 3UG4841 to use with S7-300/400 controllers! / IO-Link Geraete FB fuer SIRIUS 3UG4841 zur Nutzung mit S7-1500!
   VAR_INPUT
      execute : Bool;   // Request to execute function / Auftrag starten (mit steigender Flanke)
      logicalAddr : DInt;   // Logical address of IO-Link master module (sub module for ET 200eco PN) / Logische EA-Adresse des IO-Link Master Moduls
      cap : Int := 227;   // Client Access Point; 0xB400 for ET 200eco PN, CM 8x IO-Link, else 0xE003 (227) / Client Access Point (CAP), Siemens IO-Link Master immer 227 dezimal
      readWrite : Bool;   // FALSE: read, TRUE: write / Lese-/Schreibzugriff: 0=Lesen, 1=Schreiben
      port : Int;   // Port of the IO-Link Master for the Device / Port des Geraetes am IO-Link Mastermodul
      parameterPage0 : Bool;   // Read access on parameter page 0 / Lesen Parameter Page 0
      systemCommands : Bool;   // Write system commands / Schreiben Systemkommandos
      vendorName : Bool;   // Read vendor name / Lesen Herstellername
      vendorText : Bool;   // Read vendor text / Lesen Herstellertext
      productName : Bool;   // Read product name / Lesen Produktname
      productID : Bool;   // Read product ID / Lesen Produkt ID
      hwRevision : Bool;   // Read hardware revision / Lesen HW-Revision
      fwRevision : Bool;   // Read firmware revision / Lesen FW-Revision
      appSpecificName : Bool;   // Read/Write application specific name / Lesen/Schreiben des spezifischen Applikationsnamen
      diagnostics : Bool;   // Read diagnostics / Lesen der Diagnose
      measurements : Bool;   // Read measurements / Lesen der Messwerte
      parameters : Bool;   // Read/Write parameters / Lesen/Schreiben der Parameter
   END_VAR
   VAR_OUTPUT
      done : Bool;   // TRUE: Commanded functionality has been completed successfully / Gueltigkeit 0: Daten ungueltig ; 1: Daten gueltig
      busy : Bool;   // TRUE: FB is not finished and new output values can be expected / 0: Auftrag beendet 1: Auftrag in Bearbeitung
      error : Bool;   // TRUE: An error occurred during the execution of the FB / Fehler = 0: kein Fehler; 1: Funktionsabbruch mit Fehler
      status : Word;   // 16#0000 - 16#7FFF: Status of the FB, 16#8000 - 16#FFFF: Error identification / DP/ PNIO - Fehlerstatus ; ERROR = 1 - Kommunikationsfehler in Detail
      diagDeviceFB : "LIOLink_typeDiagnostics";   // Diagnostics information of LIOLink_Device / IO-Link - Fehlerstatus; ERROR = 1: IO-Link Fehler in Detail
   END_VAR
   VAR_IN_OUT
      data : "LIOLink_3UG4841_typeAll";   // Data area, device specific (Data Type) / Ablage der Gerätedaten, gerätespezifisch (Datentyp in DB)
   END_VAR
   VAR
      instDevice : "LIOLink_Device";
      statRecordParam : Struct   // Parameters to read/write specific records / Datensatzparameter (geraetespezifisch)
         index : Array[0..28] of Int;   // Index of data set / Datensatzindex
         subindex : Array[0..28] of Int;   // Subindex of data sets / Datensatzsubindex
         length : Array[0..28] of Int;   // Length of data set / Datensatzlänge
      END_STRUCT;
      statRecord : Array[0..231] of Byte;   // Record buffer
      statParameterPage0 AT statRecord : "LIOLink_typeParameterPage0";
      statVendorName AT statRecord : String[11];
      statVendorText AT statRecord : String[64];
      statProductName AT statRecord : String[64];
      statProductID AT statRecord : String[14];
      statHWRevision AT statRecord : String[7];
      statFWRevision AT statRecord : String[7];
      statAppSpecName AT statRecord : String[32];
      statDiagnostics AT statRecord : "LIOLink_3UG4841_typeDiag";
      statMeasurements AT statRecord : "LIOLink_3UG4841_typeMeasure";
      statParameters AT statRecord : "LIOLink_3UG4841_typeParam";   // Product family SIRIUS (0x60)
      statSystemCommands AT statRecord : Byte;
      statIndex : Int;   // Requested index
      statSubindex : Int;   // Requested subindex
      statRecordLen : Int;   // Length of record to be written
      statRequest : Int;   // Case of request (data set) / Aktueller Fall (anfgefragter Datensatz)
      statDoneOld : Bool;   // Last cycle's value of instDevice.done
   END_VAR
   VAR_TEMP
      tempIndex : Int;   // Loop index
      tempLen : Int;   // Length
   END_VAR
   VAR CONSTANT
      MODE_READ : Bool := FALSE;   // Mode to read data
      MODE_WRITE : Bool := TRUE;   // Mode to write data
      STATUS_IDLE : Word := 16#7000;   // Status: Idle
   END_VAR
   // statRecordParam.index[3] := 2;
   // statRecordParam.index[2] := 0;
   // statRecordParam.index[1] := 0;
   // statRecordParam.index[0] := 0;
   // statRecordParam.index[17] := 23;
   // statRecordParam.index[16] := 22;
   // statRecordParam.index[5] := 0;
   // statRecordParam.index[4] := 0;
   // statRecordParam.index[15] := 21;
   // statRecordParam.index[14] := 20;
   // statRecordParam.index[13] := 19;
   // statRecordParam.index[12] := 18;
   // statRecordParam.index[11] := 17;
   // statRecordParam.index[10] := 16;
   // statRecordParam.index[9] := 0;
   // statRecordParam.index[8] := 0;
   // statRecordParam.index[7] := 0;
   // statRecordParam.index[6] := 0;
   // statRecordParam.length[28] := 74;
   // statRecordParam.length[27] := 0;
   // statRecordParam.length[26] := 0;
   // statRecordParam.length[25] := 50;
   // statRecordParam.length[24] := 30;
   // statRecordParam.length[23] := 0;
   // statRecordParam.length[22] := 0;
   // statRecordParam.length[21] := 0;
   // statRecordParam.length[20] := 0;
   // statRecordParam.length[19] := 0;
   // statRecordParam.length[18] := 32;
   // statRecordParam.length[17] := 7;
   // statRecordParam.length[16] := 7;
   // statRecordParam.length[15] := 0;
   // statRecordParam.length[14] := 0;
   // statRecordParam.length[13] := 14;
   // statRecordParam.length[12] := 64;
   // statRecordParam.length[11] := 64;
   // statRecordParam.length[10] := 11;
   // statRecordParam.length[9] := 0;
   // statRecordParam.length[8] := 0;
   // statRecordParam.length[7] := 0;
   // statRecordParam.length[6] := 0;
   // statRecordParam.length[5] := 0;
   // statRecordParam.length[4] := 0;
   // statRecordParam.length[3] := 1;
   // statRecordParam.length[2] := 0;
   // statRecordParam.length[1] := 16;
   // statRecordParam.length[0] := 0;
   // statRecordParam.index[28] := 131;
   // statRecordParam.index[27] := 0;
   // statRecordParam.index[26] := 0;
   // statRecordParam.index[25] := 94;
   // statRecordParam.index[24] := 92;
   // statRecordParam.index[23] := 0;
   // statRecordParam.index[22] := 0;
   // statRecordParam.index[21] := 0;
   // statRecordParam.index[20] := 0;
   // statRecordParam.index[19] := 0;
   // statRecordParam.index[18] := 24;
BEGIN
   REGION BLOCK INFO HEADER
     //===============================================================================
     // Siemens / (c)Copyright 2020
     //-------------------------------------------------------------------------------
     // Title:            LIOLink_3UG4841
     // Function:         Capsule block to communicate with 3UG4841 devices
     // Library:          LIOLink
     // Author:           Siemens Industry Online Support
     // Tested with:      CPU 317-2 PN/DP FW 3.2
     // Engineering:      TIA Portal V16
     // Restrictions:     --
     // Requirements:     --
     //-------------------------------------------------------------------------------
     // Change log table:
     // Version  | Date       | Expert in charge       | Changes applied
     //----------|------------|------------------------|------------------------------
     // 01.00.00 | 11.04.2014 | Online Support         | First release
     // 01.01.00 | 12.09.2014 | Online Support         | Bugfixing write case 28 (data set 131)
     // 02.00.00 | 30.03.2015 | Online Support         | Upgrade to TIA Portal V13 SP1, use function IO_LINK_DEVICE, only one function for S7-1200 and 1500
     // 02.01.00 | 23.10.2015 | Online Support         | Upgraded FB "IO_LINK_DEVICE to V3.1.0
     // 03.00.00 | 22.09.2020 | Online Support         | Rewrote block for FB "LIOLink_Device" V4.0.0
     //===============================================================================
   END_REGION

   REGION INIT
     IF (#execute = TRUE AND #instDevice.status = #STATUS_IDLE) THEN
       // Request selector
       IF #parameterPage0 THEN
         #statRequest := 1;
       ELSIF #systemCommands THEN
         #statRequest := 3;
       ELSIF #vendorName THEN
         #statRequest := 10;
       ELSIF #vendorText THEN
         #statRequest := 11;
       ELSIF #productName THEN
         #statRequest := 12;
       ELSIF #productID THEN
         #statRequest := 13;
       ELSIF #hwRevision THEN
         #statRequest := 16;
       ELSIF #fwRevision THEN
         #statRequest := 17;
       ELSIF #appSpecificName THEN
         #statRequest := 18;
       ELSIF #diagnostics THEN
         #statRequest := 24;
       ELSIF #measurements THEN
         #statRequest := 25;
       ELSIF #parameters THEN
         #statRequest := 28;
       ELSE
         #statRequest := 0;
       END_IF;

       // Set request specific parameters
       #statIndex := #statRecordParam.index[#statRequest];
       #statSubindex := #statRecordParam.subindex[#statRequest];
       #statRecordLen := #statRecordParam.length[#statRequest];

       IF #readWrite = #MODE_WRITE THEN
         REGION write
           CASE #statRequest OF
             3:
               #statSystemCommands := #data.systemCommands;
             18:
               #statAppSpecName := #data.appSpecificName; // copy text into writing data
               #tempLen := LEN(#statAppSpecName); // determine length of text

               // Shift chars in array to remove String header
               FOR #tempIndex := 0 TO #tempLen - 1 DO
                 #statRecord[#tempIndex] := #statRecord[#tempIndex + 2]; // move [2] to [0], [3] to [1] ... until end of String
               END_FOR;

               // Fill remaining characters with null
               FOR #tempIndex := #tempLen TO #statRecordLen - 1 DO
                 #statRecord[#tempIndex] := CHAR_TO_BYTE('$00');
               END_FOR;
             28:
               #statParameters := #data.parameters;
             ELSE // All other data sets are read only  
               ;
           END_CASE;
         END_REGION

       END_IF;
     END_IF;
   END_REGION

   REGION CALL
     #instDevice(execute     := #execute,
                 logicalAddr := #logicalAddr,
                 cap         := #cap,
                 readWrite   := #readWrite,
                 "port"      := #port,
                 index       := #statIndex,
                 subindex    := #statSubindex,
                 writeLen    := #statRecordLen,
                 timeout     := T#20s,
                 record      := #statRecord);
   END_REGION

   REGION READ
     // Copy data
     IF #instDevice.done = TRUE AND #statDoneOld = FALSE AND #readWrite = #MODE_READ THEN
       IF (#statRequest >= 10 AND #statRequest <= 18) THEN // Only applies for String parameters (case 10..18)
         // Shift all characters to add string header
         FOR #tempIndex := (#statRecordLen + 1) TO 2 BY -1 DO
           #statRecord[#tempIndex] := #statRecord[#tempIndex - 2];
         END_FOR;
         // Add String header
         #statRecord[0] := INT_TO_BYTE(#statRecordLen);
         #statRecord[1] := INT_TO_BYTE(#statRecordLen);
       END_IF;

       CASE #statRequest OF
         1:
           #data.parameterPage0 := #statParameterPage0;
         10:
           #data.vendorName := #statVendorName;
         11:
           #data.vendorText := #statVendorText;
         12:
           #data.productName := #statProductName;
         13:
           #data.productID := #statProductID;
         16:
           #data.hwRevision := #statHWRevision;
         17:
           #data.fwRevision := #statFWRevision;
         18:
           #data.appSpecificName := #statAppSpecName;
         24:
           #data.diagnostics := #statDiagnostics;
         25:
           #data.measuredValues := #statMeasurements;
         28:
           #data.parameters := #statParameters;
         ELSE // Other data sets are not defined
           ;
       END_CASE;
     END_IF;

     #statDoneOld := #instDevice.done;
   END_REGION

   REGION OUTPUTS
     #done := #instDevice.done;
     #busy := #instDevice.busy;
     #error := #instDevice.error;
     #status := #instDevice.status;
     #diagDeviceFB := #instDevice.diagnostics;
   END_REGION
END_FUNCTION_BLOCK

FUNCTION_BLOCK "LIOLink_3UG4851"   // FB5190, SCL
TITLE = LIOLink_3UG4851 / IO_LINK_3UG4851_1500
{ S7_Optimized_Access := 'FALSE' }
AUTHOR : SIOS
FAMILY : LIOLink
VERSION : 3.0
// IO-Link Device FB for SIRIUS 3UG4851 to use with S7-300/400 controllers! / IO-Link Geraete FB fuer SIRIUS 3UG4851 zur Nutzung mit S7-1500!
   VAR_INPUT
      execute : Bool;   // Request to execute function / Auftrag starten (mit steigender Flanke)
      logicalAddr : DInt;   // Logical address of IO-Link master module (sub module for ET 200eco PN) / Logische EA-Adresse des IO-Link Master Moduls
      cap : Int := 227;   // Client Access Point; 0xB400 for ET 200eco PN, CM 8x IO-Link, else 0xE003 (227) / Client Access Point (CAP), Siemens IO-Link Master immer 227 dezimal
      readWrite : Bool;   // FALSE: read, TRUE: write / Lese-/Schreibzugriff: 0=Lesen, 1=Schreiben
      port : Int;   // Port of the IO-Link Master for the Device / Port des Geraetes am IO-Link Mastermodul
      parameterPage0 : Bool;   // Read access on parameter page 0 / Lesen Parameter Page 0
      systemCommands : Bool;   // Write system commands / Schreiben Systemkommandos
      vendorName : Bool;   // Read vendor name / Lesen Herstellername
      vendorText : Bool;   // Read vendor text / Lesen Herstellertext
      productName : Bool;   // Read product name / Lesen Produktname
      productID : Bool;   // Read product ID / Lesen Produkt ID
      hwRevision : Bool;   // Read hardware revision / Lesen HW-Revision
      fwRevision : Bool;   // Read firmware revision / Lesen FW-Revision
      appSpecificName : Bool;   // Read/Write application specific name / Lesen/Schreiben des spezifischen Applikationsnamen
      diagnostics : Bool;   // Read diagnostics / Lesen der Diagnose
      measurements : Bool;   // Read measurements / Lesen der Messwerte
      parameters : Bool;   // Read/Write parameters / Lesen/Schreiben der Parameter
   END_VAR
   VAR_OUTPUT
      done : Bool;   // TRUE: Commanded functionality has been completed successfully / Gueltigkeit 0: Daten ungueltig ; 1: Daten gueltig
      busy : Bool;   // TRUE: FB is not finished and new output values can be expected / 0: Auftrag beendet 1: Auftrag in Bearbeitung
      error : Bool;   // TRUE: An error occurred during the execution of the FB / Fehler = 0: kein Fehler; 1: Funktionsabbruch mit Fehler
      status : Word;   // 16#0000 - 16#7FFF: Status of the FB, 16#8000 - 16#FFFF: Error identification / DP/ PNIO - Fehlerstatus ; ERROR = 1 - Kommunikationsfehler in Detail
      diagDeviceFB : "LIOLink_typeDiagnostics";   // Diagnostics information of LIOLink_Device / IO-Link - Fehlerstatus; ERROR = 1: IO-Link Fehler in Detail
   END_VAR
   VAR_IN_OUT
      data : "LIOLink_3UG4851_typeAll";   // Data area, device specific (Data Type) / Ablage der Gerätedaten, gerätespezifisch (Datentyp in DB)
   END_VAR
   VAR
      instDevice : "LIOLink_Device";
      statRecordParam : Struct   // Parameters to read/write specific records / Datensatzparameter (geraetespezifisch)
         index : Array[0..28] of Int;   // Index of data set / Datensatzindex
         subindex : Array[0..28] of Int;   // Subindex of data sets / Datensatzsubindex
         length : Array[0..28] of Int;   // Length of data set / Datensatzlänge
      END_STRUCT;
      statRecord : Array[0..231] of Byte;   // Record buffer
      statParameterPage0 AT statRecord : "LIOLink_typeParameterPage0";
      statVendorName AT statRecord : String[11];
      statVendorText AT statRecord : String[64];
      statProductName AT statRecord : String[64];
      statProductID AT statRecord : String[14];
      statHWRevision AT statRecord : String[7];
      statFWRevision AT statRecord : String[7];
      statAppSpecName AT statRecord : String[32];
      statDiagnostics AT statRecord : "LIOLink_3UG4851_typeDiag";
      statMeasurements AT statRecord : "LIOLink_3UG4851_typeMeasure";
      statParameters AT statRecord : "LIOLink_3UG4851_typeParam";   // Product family SIRIUS (0x60)
      statSystemCommands AT statRecord : Byte;
      statIndex : Int;   // Requested index
      statSubindex : Int;   // Requested subindex
      statRecordLen : Int;   // Length of record to be written
      statRequest : Int;   // Case of request (data set) / Aktueller Fall (anfgefragter Datensatz)
      statDoneOld : Bool;   // Last cycle's value of instDevice.done
   END_VAR
   VAR_TEMP
      tempIndex : Int;   // Loop index
      tempLen : Int;   // Length
   END_VAR
   VAR CONSTANT
      MODE_READ : Bool := FALSE;   // Mode to read data
      MODE_WRITE : Bool := TRUE;   // Mode to write data
      STATUS_IDLE : Word := 16#7000;   // Status: Idle
   END_VAR
   // statRecordParam.index[3] := 2;
   // statRecordParam.index[2] := 0;
   // statRecordParam.index[1] := 0;
   // statRecordParam.index[0] := 0;
   // statRecordParam.index[17] := 23;
   // statRecordParam.index[16] := 22;
   // statRecordParam.index[5] := 0;
   // statRecordParam.index[4] := 0;
   // statRecordParam.index[15] := 21;
   // statRecordParam.index[14] := 20;
   // statRecordParam.index[13] := 19;
   // statRecordParam.index[12] := 18;
   // statRecordParam.index[11] := 17;
   // statRecordParam.index[10] := 16;
   // statRecordParam.index[9] := 0;
   // statRecordParam.index[8] := 0;
   // statRecordParam.index[7] := 0;
   // statRecordParam.index[6] := 0;
   // statRecordParam.length[28] := 48;
   // statRecordParam.length[27] := 0;
   // statRecordParam.length[26] := 0;
   // statRecordParam.length[25] := 18;
   // statRecordParam.length[24] := 30;
   // statRecordParam.length[23] := 0;
   // statRecordParam.length[22] := 0;
   // statRecordParam.length[21] := 0;
   // statRecordParam.length[20] := 0;
   // statRecordParam.length[19] := 0;
   // statRecordParam.length[18] := 32;
   // statRecordParam.length[17] := 7;
   // statRecordParam.length[16] := 7;
   // statRecordParam.length[15] := 0;
   // statRecordParam.length[14] := 0;
   // statRecordParam.length[13] := 14;
   // statRecordParam.length[12] := 64;
   // statRecordParam.length[11] := 64;
   // statRecordParam.length[10] := 11;
   // statRecordParam.length[9] := 0;
   // statRecordParam.length[8] := 0;
   // statRecordParam.length[7] := 0;
   // statRecordParam.length[6] := 0;
   // statRecordParam.length[5] := 0;
   // statRecordParam.length[4] := 0;
   // statRecordParam.length[3] := 1;
   // statRecordParam.length[2] := 0;
   // statRecordParam.length[1] := 16;
   // statRecordParam.length[0] := 0;
   // statRecordParam.index[28] := 131;
   // statRecordParam.index[27] := 0;
   // statRecordParam.index[26] := 0;
   // statRecordParam.index[25] := 94;
   // statRecordParam.index[24] := 92;
   // statRecordParam.index[23] := 0;
   // statRecordParam.index[22] := 0;
   // statRecordParam.index[21] := 0;
   // statRecordParam.index[20] := 0;
   // statRecordParam.index[19] := 0;
   // statRecordParam.index[18] := 24;
BEGIN
   REGION BLOCK INFO HEADER
     //===============================================================================
     // Siemens / (c)Copyright 2020
     //-------------------------------------------------------------------------------
     // Title:            LIOLink_3UG4851
     // Function:         Capsule block to communicate with 3UG4851 devices
     // Library:          LIOLink
     // Author:           Siemens Industry Online Support
     // Tested with:      CPU 317-2 PN/DP FW 3.2
     // Engineering:      TIA Portal V16
     // Restrictions:     --
     // Requirements:     --
     //-------------------------------------------------------------------------------
     // Change log table:
     // Version  | Date       | Expert in charge       | Changes applied
     //----------|------------|------------------------|------------------------------
     // 01.00.00 | 11.04.2014 | Online Support         | First release
     // 01.01.00 | 12.09.2014 | Online Support         | Bugfixing write case 28 (data set 131)
     // 02.00.00 | 30.03.2015 | Online Support         | Upgrade to TIA Portal V13 SP1, use function IO_LINK_DEVICE, only one function for S7-1200 and 1500
     // 02.01.00 | 23.10.2015 | Online Support         | Upgraded FB "IO_LINK_DEVICE to V3.1.0
     // 03.00.00 | 22.09.2020 | Online Support         | Rewrote block for FB "LIOLink_Device" V4.0.0
     //===============================================================================
   END_REGION

   REGION INIT
     IF (#execute = TRUE AND #instDevice.status = #STATUS_IDLE) THEN
       // Request selector
       IF #parameterPage0 THEN
         #statRequest := 1;
       ELSIF #systemCommands THEN
         #statRequest := 3;
       ELSIF #vendorName THEN
         #statRequest := 10;
       ELSIF #vendorText THEN
         #statRequest := 11;
       ELSIF #productName THEN
         #statRequest := 12;
       ELSIF #productID THEN
         #statRequest := 13;
       ELSIF #hwRevision THEN
         #statRequest := 16;
       ELSIF #fwRevision THEN
         #statRequest := 17;
       ELSIF #appSpecificName THEN
         #statRequest := 18;
       ELSIF #diagnostics THEN
         #statRequest := 24;
       ELSIF #measurements THEN
         #statRequest := 25;
       ELSIF #parameters THEN
         #statRequest := 28;
       ELSE
         #statRequest := 0;
       END_IF;

       // Set request specific parameters
       #statIndex := #statRecordParam.index[#statRequest];
       #statSubindex := #statRecordParam.subindex[#statRequest];
       #statRecordLen := #statRecordParam.length[#statRequest];

       IF #readWrite = #MODE_WRITE THEN
         REGION write
           CASE #statRequest OF
             3:
               #statSystemCommands := #data.systemCommands;
             18:
               #statAppSpecName := #data.appSpecificName; // copy text into writing data
               #tempLen := LEN(#statAppSpecName); // determine length of text

               // Shift chars in array to remove String header
               FOR #tempIndex := 0 TO #tempLen - 1 DO
                 #statRecord[#tempIndex] := #statRecord[#tempIndex + 2]; // move [2] to [0], [3] to [1] ... until end of String
               END_FOR;

               // Fill remaining characters with null
               FOR #tempIndex := #tempLen TO #statRecordLen - 1 DO
                 #statRecord[#tempIndex] := CHAR_TO_BYTE('$00');
               END_FOR;
             28:
               #statParameters := #data.parameters;
             ELSE // All other data sets are read only  
               ;
           END_CASE;
         END_REGION

       END_IF;
     END_IF;
   END_REGION

   REGION CALL
     #instDevice(execute     := #execute,
                 logicalAddr := #logicalAddr,
                 cap         := #cap,
                 readWrite   := #readWrite,
                 "port"      := #port,
                 index       := #statIndex,
                 subindex    := #statSubindex,
                 writeLen    := #statRecordLen,
                 timeout     := T#20s,
                 record      := #statRecord);
   END_REGION

   REGION READ
     // Copy data
     IF #instDevice.done = TRUE AND #statDoneOld = FALSE AND #readWrite = #MODE_READ THEN
       IF (#statRequest >= 10 AND #statRequest <= 18) THEN // Only applies for String parameters (case 10..18)
         // Shift all characters to add string header
         FOR #tempIndex := (#statRecordLen + 1) TO 2 BY -1 DO
           #statRecord[#tempIndex] := #statRecord[#tempIndex - 2];
         END_FOR;
         // Add String header
         #statRecord[0] := INT_TO_BYTE(#statRecordLen);
         #statRecord[1] := INT_TO_BYTE(#statRecordLen);
       END_IF;

       CASE #statRequest OF
         1:
           #data.parameterPage0 := #statParameterPage0;
         10:
           #data.vendorName := #statVendorName;
         11:
           #data.vendorText := #statVendorText;
         12:
           #data.productName := #statProductName;
         13:
           #data.productID := #statProductID;
         16:
           #data.hwRevision := #statHWRevision;
         17:
           #data.fwRevision := #statFWRevision;
         18:
           #data.appSpecificName := #statAppSpecName;
         24:
           #data.diagnostics := #statDiagnostics;
         25:
           #data.measuredValues := #statMeasurements;
         28:
           #data.parameters := #statParameters;
         ELSE // Other data sets are not defined
           ;
       END_CASE;
     END_IF;

     #statDoneOld := #instDevice.done;
   END_REGION

   REGION OUTPUTS
     #done := #instDevice.done;
     #busy := #instDevice.busy;
     #error := #instDevice.error;
     #status := #instDevice.status;
     #diagDeviceFB := #instDevice.diagnostics;
   END_REGION
END_FUNCTION_BLOCK

// folder: Devices/SIMATIC RF200

FUNCTION_BLOCK "LIOLink_RF200_ReadTag"   // FB2, SCL
TITLE = LRfidIOL_Read
{ S7_Optimized_Access := 'FALSE' }
FAMILY : S7-300
VERSION : 3.1
// Read Data with IO-Link readers
// IO-Link V1.1
   VAR_INPUT
      execute : Bool;
      addrTag : Word;
      length : Word;
      hwID : Word;
      portAddr : Int;
      "version" : Int;
   END_VAR
   VAR_OUTPUT
      done : Bool;
      busy : Bool;
      error : Bool;
      status : DWord;
      statusWord AT status : Array[0..1] of Word;
      presence : Bool;
   END_VAR
   VAR_IN_OUT
      identData : ANY;
   END_VAR
   VAR
      statPae : Array[0..28] of Byte;
      Status_Byte : Byte;
      Status_bit AT Status_Byte : Array[0..7] of Bool;
      statPresence : Bool;
      statNState : Int;
      statIdleState : Int;
      statTelegramState : Int := 1;
      statReadState : Int := 2;
      statErrorState : Int := 3;
      statAdr : Word;
      statAdrRead AT statAdr : Array[0..1] of Byte;
      statBlk : Int;
      statReadOffset : Int := 0;
      statExecuteReq : Bool;
      statOffset : DInt;
      statOffset2 : DWord;
      statLength : DInt;
      statDat : Array[0..31] of Byte;
      statRecDat : Array[0..31] of Byte;
      statAddrOffset : Int;
      statPresenceFF : Bool;
      statTimerIn : Bool;
      statTimerPt : Time := T#5s;
      instTon : TON;
      statDone : Bool;
      statBusy : Bool;
      InstSetIoPart : SETIO_PART;
      statIoPartError : Bool;
      statIoPartStatus : DWord;
      InstGetIoPart : GETIO_PART;
      statIOsizeNetto : Int;
      statIOsize : Int;
   END_VAR
   VAR_TEMP
      tempSPointer : ANY;
      tempPoint1 AT tempSPointer : Struct
         dentifier : Byte;
         typ : Byte;
         length : Int;
         dbnr : Int;
         datapointer : DWord;
      END_STRUCT;
      tempDPointer : ANY;
      tempPoint2 AT tempDPointer : Struct
         dentifier : Byte;
         typ : Byte;
         length : Int;
         dbnr : Int;
         datapointer : DWord;
      END_STRUCT;
      tempError : Bool;
      tempStatus : DWord;
      tempStatusWord AT tempStatus : Array[0..1] of Word;
   END_VAR
   VAR CONSTANT
      VERSION_10 : Int := 10;   // Identifier IO-Link version 1.0
      VERSION_11 : Int := 11;   // Identifier IO-Link version 1.1
      IOL_V10 : Int := 8;
      IOL_V11 : Int := 32;
   END_VAR
BEGIN
   REGION BLOCK INFO HEADER
       //===============================================================================
       // Siemens / (c)Copyright 2020
       //-------------------------------------------------------------------------------
       // Title:            LIOLink_RF200_ReadTag
       // Function:         Reads tags from SIMATIC RF200 readers via IO-Link
       // Library:          LIOLink
       // Author:           Siemens Industry Online Support
       // Tested with:      CPU 317-2 PN/DP FW 3.2
       // Engineering:      TIA Portal V16
       // Restrictions:     --
       // Requirements:     --
       //-------------------------------------------------------------------------------
       // Change log table:
       // Version  | Date       | Expert in charge       | Changes applied
       //----------|------------|------------------------|------------------------------
       // 01.00.00 | 01.07.2013 | Online Support         | First release
       // 01.01.00 | 01.12.2016 | Online Support         | Upgrade to TIA Portal V14
       // 02.00.00 | 01.09.2017 | Online Support         | Upgrade to TIA Portal V14 SP1
       //                                                | Implementation of Programming styleguide
       //                                                | Added support for IO-Link V1.1 readers
       // 02.01.00 | 01.12.2017 | Online Support         | Bug fixes and performance improvements
       // 02.02.00 | 01.03.2020 | Online Support         | Upgrade to TIA Portal V16
       // 02.03.00 | 08.03.2020 | Online Support         | Added input "version" for IO-Link version / bug fix  
       //===============================================================================
   END_REGION

   IF #version = #VERSION_11 THEN                               //determine IO-Link reader version (1.0/1.1) to set offsets
       #statIOsize := #IOL_V11;
       #statIOsizeNetto := #IOL_V11 - 4;
   ELSE
       #statIOsize := #IOL_V10;
       #statIOsizeNetto := #IOL_V10 - 4;
   END_IF;

   #statAddrOffset:=#portAddr;                           //start adress of port
   #InstGetIoPart(ID := #hwID,
                 OFFSET := #statAddrOffset,
                 LEN := #statIOsize,
                 STATUS => #statIoPartStatus,
                 ERROR => #statIoPartError,
                 INPUTS := #statRecDat);

   #Status_Byte:=#statRecDat[0];                           //Status Byte
   #statPresence:=#Status_bit[5];                       //Presence bit. Transponder on field
   #presence:=#statPresence;

   IF NOT #execute THEN
      #statDone := false;
      #statBusy := false;
      #done := false;
      #busy := false;
      #error := false;
      #status := 0;
   ELSE
      #done := #statDone;
      #busy := #statBusy;
   END_IF;

   IF #execute AND #execute<> #statExecuteReq THEN        //Positive edge for d#reading of data
     IF NOT #statBusy THEN
       #statAdr:=#addrTag;                                 //Transpoder Adress
       #statLength:=#length;                             //Length of read Data
       #statBusy:=TRUE;
       #statDone:=FALSE;                                   //reset all the output parameters                                   
       #error:=FALSE;
       #status:=0;
       #statReadOffset:=0;
       #statNState:=#statReadState;                          //next step >> send read command
     ELSE
       #tempStatusWord[1]:=16#8102;                          //block is still active
       #tempStatusWord[0]:=16#0001;                          //Error identifier for block errors
       #status := #tempStatus;
       #statNState:=#statErrorState;
   END_IF;
   IF #statLength < #statIOsizeNetto THEN
       #tempStatusWord[1] := 16#8104;                              //length too short
       #tempStatusWord[0] := 16#0001;                              //identifier rfid errors
       #status := #tempStatus;
       #statNState := #statErrorState;
   END_IF;
   END_IF;
   #statExecuteReq:=#execute;


   IF NOT #presence AND #presence<>#statPresenceFF THEN   //the tag has left the antenna  field
       IF NOT #statDone THEN
       #statTimerIn:=true;                              //wait 5 sec
     END_IF;
   END_IF;
   #statPresenceFF:=#presence;
   IF #presence THEN
     #statTimerIn:=false;
   END_IF;
   //-----------------------------------------------------------------------------------------------------//
   //------------------------------------------start of state machine------------------------------------//
   //-----------------------------------------------------------------------------------------------------//

   CASE #statNState OF
   0://idle
     #statReadOffset:=0;                                             //offset of puffer must be reseted
     #statBusy:=false;
     #statTimerIn:=false;

   //-------------------------------------------------Read state------------------------------------------//
   //---------------------------------------------sent read command---------------------------------------//
   //-----------------------------------------------------------------------------------------------------//

   2: //READ_state

      IF #statLength>0 THEN  
          #statDat[0]:= 16#2;                      //Set read command
          #statDat[2]:=#statAdrRead[0];             //Adr_H
          #statDat[3]:=#statAdrRead[1];             //Adr-L
      END_IF;

       IF #statBlk=0 THEN
         #statNState:=#statTelegramState;                           //Telegram: Edit the read data
       END_IF;


   //-----------------------------------------------Telegram state----------------------------------------//
   //---------------------------------------------edit received data--------------------------------------//
   //-----------------------------------------------------------------------------------------------------//  

   1://Telegram

    IF #statLength>0 THEN                                  //Only when length of data > 0 can continue  
     IF #Status_bit[6] THEN                            //IF RFID error has occured
       #tempStatusWord[1]:=#statRecDat[1];          //error_RFID
       #tempStatusWord[0]:=16#0011;                          //Error identifier for RFID errors
       #status := #tempStatus;
       #statNState:=#statErrorState;
     END_IF;

   //-------------------------- read command is ready------------------------------------------------//

     IF #Status_bit[7] AND #Status_bit[1]  THEN  
       IF #statRecDat[2]=#statAdrRead[0] AND #statRecDat[3]=#statAdrRead[1] THEN //received ADR must be ==sent ADR
          #statPae[0] := #statRecDat[4];                             //Save of read data
          #statPae[1] := #statRecDat[5];
          #statPae[2] := #statRecDat[6];
          #statPae[3] := #statRecDat[7];
          #statPae[4] := #statRecDat[8];
          #statPae[5] := #statRecDat[9];
          #statPae[6] := #statRecDat[10];
          #statPae[7] := #statRecDat[11];
          #statPae[8] := #statRecDat[12];
          #statPae[9] := #statRecDat[13];
          #statPae[10] := #statRecDat[14];
          #statPae[11] := #statRecDat[15];
          #statPae[12] := #statRecDat[16];
          #statPae[13] := #statRecDat[17];
          #statPae[14] := #statRecDat[18];
          #statPae[15] := #statRecDat[19];
          #statPae[16] := #statRecDat[20];
          #statPae[17] := #statRecDat[21];
          #statPae[18] := #statRecDat[22];
          #statPae[19] := #statRecDat[23];
          #statPae[20] := #statRecDat[24];
          #statPae[21] := #statRecDat[25];
          #statPae[22] := #statRecDat[26];
          #statPae[23] := #statRecDat[27];
          #statPae[24] := #statRecDat[28];
          #statPae[25] := #statRecDat[29];
          #statPae[26] := #statRecDat[30];
          #statPae[27] := #statRecDat[31];

          #tempSPointer:=#statPae[0];
          #tempDPointer:=#identData;                             //Destination pointer
          #statOffset:=DWORD_TO_DINT(#tempPoint2.datapointer);  //offset of destination pointer
          #statOffset2:=DINT_TO_DWORD(#statOffset/8+#statReadOffset);
          #statOffset2:=16#84000000 OR SHL(IN:=#statOffset2, N:=3);
          #tempPoint2.datapointer:=#statOffset2;               //Offset of data block
          IF #statLength >= #statIOsizeNetto THEN
              #tempPoint1.length := #statIOsizeNetto;                        //length of data, that must be saved                       
              #tempPoint2.length := #statIOsizeNetto;
          ELSIF #statLength > 0 AND #statLength < #statIOsizeNetto THEN
              #tempPoint1.length := DINT_TO_INT(#statLength);
              #tempPoint2.length := DINT_TO_INT(#statLength);
          END_IF;

          #statBlk:=BLKMOV(SRCBLK:=#tempSPointer, DSTBLK=>#tempDPointer); //Copy the read Data into the data block-buffer

         IF #statBlk=0 THEN

              IF #Status_bit[7] AND NOT #Status_bit[6] THEN
                  #statLength:=#statLength-#statIOsizeNetto;
                  #statReadOffset:=#statReadOffset+#statIOsizeNetto;                                   //offset must be changed
                   #statAdr:=INT_TO_WORD(WORD_TO_INT(#statAdr) + #statIOsizeNetto);     //Change the ADR (#statIOsizeNetto Bytes)       
                #statNState:=#statReadState;                      //Start a new read command
            ELSE
                #statNState:=#statIdleState;
              END_IF;
          ELSE
            #tempStatusWord[1]:=INT_TO_WORD(#statBlk);                 //Error has to BLKMOV occured
            #tempStatusWord[0]:=16#0001;                           //functions-Error identifier
            #status := #tempStatus;
            #statNState:=#statErrorState;
          END_IF;
        END_IF;
       END_IF; 

   ELSE
      #statNState := #statIdleState;
      #statBusy := FALSE;
      #statDone := TRUE;
      #done := TRUE;
      #busy := FALSE;

      #statDat[0] := 16#0;                                          //Reset read command
      #InstSetIoPart(ID      := #hwID,
                     OFFSET  := #statAddrOffset,
                     LEN     := #statIOsize,
                     STATUS  => #statIoPartStatus,
                     ERROR   => #statIoPartError,
                     OUTPUTS := #statDat);
   END_IF ;

   #InstSetIoPart(ID := #hwID,
                  OFFSET := #statAddrOffset,
                  LEN := #statIOsize,
                  STATUS => #statIoPartStatus,
                  ERROR => #statIoPartError,
                  OUTPUTS := #statDat);

   //------------------------------------------------------------------------------------------------------------//
   //-------------------------------------------------Error state------------------------------------------------//
   //---------------------------------------------error has occured----------------------------------------------//

   3://error
       #tempError := true;
       #error:=#tempError;
       #statBusy:=false;
       #statDone := false;
       #statTimerIn:=false;
       #statNState:=#statIdleState;

       #statDat[0] := 16#0;                                          //Reset read command
       #InstSetIoPart(ID      := #hwID,
                      OFFSET  := #statAddrOffset,
                      LEN     := #statIOsize,
                      STATUS  => #statIoPartStatus,
                      ERROR   => #statIoPartError,
                      OUTPUTS := #statDat);
   END_CASE;


   //------------------------------------------------------------------------------------------------------------//
   //-------------------------------------------------Timer------------------------------------------------------//
   //------------------------------------------------------------------------------------------------------------//


   #instTon(IN:=#statTimerIn,
                           PT:=#statTimerPt);

   IF #instTon.Q THEN                      //error has occured. No tag on field during the 5 sec.
      #tempStatusWord[1]:=16#8101;                              //tag has left the field
      #tempStatusWord[0]:=16#0001;                              //identifier rfid errors
      #status := #tempStatus;
      #statNState:=#statErrorState;
   END_IF;
END_FUNCTION_BLOCK

FUNCTION_BLOCK "LIOLink_RF200_WriteTag"   // FB3, SCL
TITLE = LRfidIOL_Write
{ S7_Optimized_Access := 'FALSE' }
FAMILY : S7-300
VERSION : 3.1
// Write Data with IO-Link readers
// IO-Link V1.1
   VAR_INPUT
      execute : Bool;
      addrTag : Word;
      length : Word;
      hwID : Word;
      portAddr : Int;
      "version" : Int;
   END_VAR
   VAR_OUTPUT
      done : Bool;
      busy : Bool;
      error : Bool;
      status : DWord;
      statusWord AT status : Array[0..1] of Word;
      presence : Bool;
   END_VAR
   VAR_IN_OUT
      identData : ANY;
   END_VAR
   VAR
      statStatusByte : Byte;
      statStatusBits AT statStatusByte : Array[0..7] of Bool;
      statPresence : Bool;
      statNState : Int;
      statIdleState : Int;
      statTelegramState : Int := 1;
      statWriteState : Int := 2;
      statErrorState : Int := 3;
      statAddr : Word;
      statAddrWrite AT statAddr : Array[0..1] of Byte;
      statBlk : Int;
      statWriteOffset : Int := 0;
      statExecuteReq : Bool;
      statLength : DInt;
      statDat : Array[0..31] of Byte;
      statRecDat : Array[0..31] of Byte;
      statAddrOffset : Int;
      statPresenceFf : Bool;
      statTImerIn : Bool;
      statTimerPT : Time := T#5s;
      instTon : TON;
      statWriteData : Array[0..1999] of Byte;
      statDiffToIOsizeNetto : Int;
      statByteMove : Int;
      statBusy : Bool;
      statDone : Bool;
      InstSetIoPart : SETIO_PART;
      statIoPartError : Bool;
      statIoPartStatus : DWord;
      InstGetIoPart : GETIO_PART;
      statIOsizeNetto : Int;
      statIOsize : Int;
   END_VAR
   VAR_TEMP
      tempError : Bool;
      tempStatus : DWord;
      tempStatusWord AT tempStatus : Array[0..1] of Word;
   END_VAR
   VAR CONSTANT
      VERSION_10 : Int := 10;   // Identifier IO-Link version 1.0
      VERSION_11 : Int := 11;   // Identifier IO-Link version 1.1
      IOL_V10 : Int := 8;
      IOL_V11 : Int := 32;
   END_VAR
BEGIN
   REGION BLOCK INFO HEADER
       //===============================================================================
       // Siemens / (c)Copyright 2020
       //-------------------------------------------------------------------------------
       // Title:            LIOLink_RF200_WriteTag
       // Function:         Write tags from SIMATIC RF200 readers via IO-Link
       // Library:          LIOLink
       // Author:           Siemens Industry Online Support
       // Tested with:      CPU 317-2 PN/DP FW 3.2
       // Engineering:      TIA Portal V16
       // Restrictions:     --
       // Requirements:     --
       //-------------------------------------------------------------------------------
       // Change log table:
       // Version  | Date       | Expert in charge       | Changes applied
       //----------|------------|------------------------|------------------------------
       // 01.00.00 | 01.07.2013 | Online Support         | First release
       // 01.01.00 | 01.12.2016 | Online Support         | Upgrade to TIA Portal V14
       // 02.00.00 | 01.09.2017 | Online Support         | Upgrade to TIA Portal V14 SP1
       //                                                | Implementation of Programming styleguide
       //                                                | Added support for IO-Link V1.1 readers
       // 02.01.00 | 01.12.2017 | Online Support         | Bug fixes and performance improvements
       // 02.02.00 | 01.03.2020 | Online Support         | Upgrade to TIA Portal V16
       // 02.03.00 | 08.03.2020 | Online Support         | Added input "version" for IO-Link version / bug fix  
       //===============================================================================
   END_REGION

   IF #version = #VERSION_11 THEN                               //determine IO-Link reader version (1.0/1.1) to set offsets
       #statIOsize := #IOL_V11;
       #statIOsizeNetto := #IOL_V11 - 4;
   ELSE
       #statIOsize := #IOL_V10;
       #statIOsizeNetto := #IOL_V10 - 4;
   END_IF;

   #statAddrOffset := #portAddr;                           //start adress of port
   #InstGetIoPart(ID := #hwID,                              //read data from process image
                  OFFSET := #statAddrOffset,
                  LEN := #statIOsize,
                  STATUS => #statIoPartStatus,
                  ERROR => #statIoPartError,
                  INPUTS := #statRecDat);
   #statStatusByte := #statRecDat[0];             //Status Byte
   #statPresence := #statStatusBits[5];                       //Presence bit. Transponder on field
   #presence := #statPresence;

   #statDiffToIOsizeNetto := WORD_TO_INT(#length) MOD #statIOsizeNetto;

   IF NOT #execute THEN
       #statDone := false;
       #statBusy := false;
       #done := false;
       #busy := false;
       #error := false;
       #status := 0;
   ELSE
       #done := #statDone;
       #busy := #statBusy;
   END_IF;

   IF #execute AND #execute <> #statExecuteReq THEN        //Positive edge for d#reading of data
       IF NOT #statBusy THEN

           #statAddr := #addrTag;                                 //Transpoder Adress
           #statLength := #length;                             //Length of read Data
           #statBusy := TRUE;
           #statDone := FALSE;                                   //reset all the output parameters                                   
           #error := FALSE;
           #status := 0;
           #statWriteOffset := 0;
           #statNState := #statWriteState;                          //next step >> send read command
       ELSE
           #tempStatusWord[1] := 16#8102;                          //block is still active
           #tempStatusWord[0] := 16#0001;                          //Error identifier for block errors
           #status := #tempStatus;
           #statNState := #statErrorState;
       END_IF;
       IF #statLength < #statIOsizeNetto THEN
           #tempStatusWord[1] := 16#8104;                              //length too short
           #tempStatusWord[0] := 16#0001;                              //identifier rfid errors
           #status := #tempStatus;
           #statNState := #statErrorState;
       END_IF;
   END_IF;
   #statExecuteReq := #execute;


   IF NOT #presence AND #presence <> #statPresenceFf THEN   //the tag has left the antenna  field
       IF NOT #statDone THEN
           #statTImerIn := true;                              //wait 5 sec
       END_IF;
   END_IF;
   #statPresenceFf := #presence;
   IF #presence THEN
       #statTImerIn := false;
   END_IF;
   //-----------------------------------------------------------------------------------------------------//
   //------------------------------------------start of state machine------------------------------------//
   //-----------------------------------------------------------------------------------------------------//

   CASE #statNState OF
      0://IDLE 
       #statWriteOffset := 0;                                             //offset of puffer must be reseted
       #statBusy := false;
       #statTImerIn := false;

       2://#Write_state

       IF #statLength > 0 THEN
           #statDat[0] := 16#1;                      //Set write command
           #statDat[2] := #statAddrWrite[0];             //Adr-H
           #statDat[3] := #statAddrWrite[1];             //Adr-L

